(* CODESYS project compile.project

Project tree, tasks and I/O mapping:
  PLCWinNT : CODESYS Control Win V3 x64, CODESYS, version 3.5.22.40
    application Application
      libraries: IoStandard, 3.5.22.0 (System); Standard, 3.5.22.0 (System)
      task MainTask (cyclic, interval 20 ms, priority 1) calls PLC_PRG
      program PLC_PRG [ST]
      function block FB_AgentProbeGood [ST]
*)

// PLCWinNT/Application/PLC_PRG
PROGRAM PLC_PRG
VAR
    _agent_template_alive : BOOL;
END_VAR

_agent_template_alive := TRUE;

END_PROGRAM

// PLCWinNT/Application/FB_AgentProbeGood
{attribute 'linkalways'}
FUNCTION_BLOCK FB_AgentProbeGood
VAR_INPUT
 x : BOOL;
END_VAR
VAR_OUTPUT
 y : BOOL;
END_VAR

y := x;

END_FUNCTION_BLOCK
